DATA_BLOCK "StationA"
{ S7_Optimized_Access := 'TRUE' }
VERSION : 0.1
NON_RETAIN
"FB_DeclarationUnit"
BEGIN
END_DATA_BLOCK
